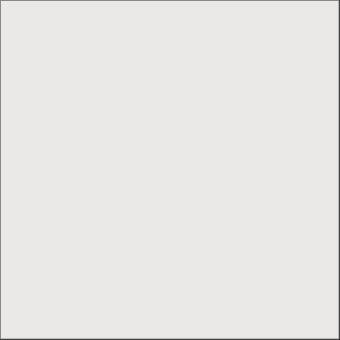
VISUALIZATION vis_InterconnectionCell  // 340x340
    Rectangle (0,0 340x340)
END_VISUALIZATION

(* stored: Version 1.1.0.1, ProductVersion 3.1.4024.12
   Visu vis_InterconnectionCell: Id {3779ae51-ab3e-4f49-a537-b5312640a47a} *)
